// TIA Portal V20 export
// export: Created 2026-10-20T18:54:47.9382926Z, ExportSetting None, DisplayName Totally Integrated Automation Portal, DisplayVersion V20 Update 6, DisplayName TIA Portal Openness, DisplayVersion V20 Update 6, DisplayName TIA Portal Version Control Interface, DisplayVersion V20 Update 6, DisplayName SINAMICS Startdrive Advanced, DisplayVersion V20 SP1, DisplayName SINAMICS Startdrive G130, G150, S120, S150, SINAMICS MV, G220, S200, S210, DisplayVersion V20 SP1, DisplayName SINAMICS Startdrive G110M, G120, G120C, G120D, G120P, G115D, DisplayVersion V20 SP1, DisplayName STEP 7 Professional, DisplayVersion V20 Update 6, DisplayName STEP 7 Safety, DisplayVersion V20 Update 2, DisplayName WinCC Basic/Comfort/Advanced, DisplayVersion V20 Update 6, DisplayName WinCC Unified, DisplayVersion V20 Update 6
VAR_GLOBAL   // PLC tag table "IO_ET200_1"
   "C1102 - SHUTTLE IN POSITION 2" AT %I107.6 : Bool;
   "C1102 - SHUTTLE IN POSITION 1" AT %I107.7 : Bool;
   "C1102 - SENSOR CNV RIGHT (PALLET DETECT 2)" AT %I107.0 : Bool;
   "C1107 - SENSOR CNV LEFT (PALLET DETECT 2)" AT %I127.1 : Bool;
   "C1107 - SHUTTLE IN POSITION 2" AT %I127.6 : Bool;
   "C1107 - SHUTTLE IN POSITION 1" AT %I127.7 : Bool;
   "C1107 - SENSOR CNV RIGHT (PALLET DETECT 2)" AT %I127.0 : Bool;
   "C1107 - SENSOR CNV RIGHT (PALLET DETECT 1)" AT %I127.5 : Bool;
   "C1102 - SENSOR CNV RIGHT (PALLET DETECT 1)" AT %I107.5 : Bool;
   "C1107 - SENSOR CNV LEFT (PALLET DETECT 1)" AT %I126.4 : Bool;
   "C1107 - SENSOR CNV LEFT" AT %I126.5 : Bool;
   "C1106 - SENSOR SAFETY PIN1 DOWN" AT %I115.3 : Bool;
   "C1107 - SENSOR SAFETY PIN1 UP" AT %I127.2 : Bool;
   "C1102 - SENSOR CNV LEFT" AT %I106.5 : Bool;
   "C1102 - SENSOR CNV LEFT (PALLET DETECT 1)" AT %I106.4 : Bool;
   "C1105 - SENSOR SAFETY PIN1 UP" AT %I113.2 : Bool;
   "C1105 - SHUTTLE IN POSITION 2" AT %I113.6 : Bool;
   "C1105 - SHUTTLE IN POSITION 1" AT %I113.7 : Bool;
   "C1105 - SENSOR CNV RIGHT (PALLET DETECT 2)" AT %I113.0 : Bool;
   "C1105 - SENSOR CNV RIGHT (PALLET DETECT 1)" AT %I113.5 : Bool;
   "C1105 - SENSOR CNV LEFT (PALLET DETECT 2)" AT %I113.1 : Bool;
   "C1105 - SENSOR CNV LEFT (PALLET DETECT 1)" AT %I112.4 : Bool;
   "C1105 - SENSOR CNV LEFT" AT %I112.5 : Bool;
   "C1104 - SENSOR SAFETY PIN1 DOWN" AT %I111.3 : Bool;
   "C1104 - SHUTTLE IN POSITION 2" AT %I111.6 : Bool;
   "C1104 - SHUTTLE IN POSITION 1" AT %I111.7 : Bool;
   "C1105 - SENSOR SAFETY PIN1 DOWN" AT %I113.3 : Bool;
   "C1104 - SENSOR CNV RIGHT (PALLET DETECT 2)" AT %I111.0 : Bool;
   "C1104 - SENSOR CNV LEFT (PALLET DETECT 2)" AT %I111.1 : Bool;
   "C1104 - SENSOR CNV LEFT (PALLET DETECT 1)" AT %I110.4 : Bool;
   "C1104 - SENSOR CNV LEFT" AT %I110.5 : Bool;
   "C1104 - SENSOR CNV RIGHT (PALLET DETECT 1)" AT %I111.5 : Bool;
   "C1106 - SENSOR CNV LEFT" AT %I114.5 : Bool;
   "C1106 - SENSOR CNV LEFT (PALLET DETECT 2)" AT %I115.1 : Bool;
   "C1106 - SENSOR CNV LEFT (PALLET DETECT 1)" AT %I114.4 : Bool;
   "C1106 - SENSOR SAFETY PIN1 UP" AT %I115.2 : Bool;
   "C1106 - SHUTTLE IN POSITION 2" AT %I115.6 : Bool;
   "C1106 - SHUTTLE IN POSITION 1" AT %I115.7 : Bool;
   "C1106 - SENSOR CNV RIGHT (PALLET DETECT 2)" AT %I115.0 : Bool;
   "C1106 - SENSOR CNV RIGHT (PALLET DETECT 1)" AT %I115.5 : Bool;
   "C1104 - SENSOR SAFETY PIN1 UP" AT %I111.2 : Bool;
   "C1102 - SENSOR CNV LEFT (PALLET DETECT 2)" AT %I107.1 : Bool;
   "C1107 - SENSOR SAFETY PIN1 DOWN" AT %I127.3 : Bool;
   "C1206 - SENSOR SAFETY PIN1 UP" AT %I345.2 : Bool;
   "C1206 - SHUTTLE IN POSITION 2" AT %I345.6 : Bool;
   "C1206 - SHUTTLE IN POSITION 1" AT %I345.7 : Bool;
   "C1206 - SENSOR CNV RIGHT (PALLET DETECT 2)" AT %I345.1 : Bool;
   "C1206 - SENSOR CNV RIGHT (PALLET DETECT 1)" AT %I344.4 : Bool;
   "C1206 - SENSOR CNV LEFT (PALLET DETECT 2)" AT %I345.0 : Bool;
   "C1206 - SENSOR CNV LEFT (PALLET DETECT 1)" AT %I345.5 : Bool;
   "C1206 - SENSOR CNV LEFT" AT %I345.4 : Bool;
   "C1205 - SENSOR SAFETY PIN1 DOWN" AT %I343.3 : Bool;
   "C1205 - SENSOR SAFETY PIN1 UP" AT %I343.2 : Bool;
   "C1205 - SENSOR CNV RIGHT (PALLET DETECT 2)" AT %I343.1 : Bool;
   "C1205 - SENSOR CNV RIGHT (PALLET DETECT 1)" AT %I342.4 : Bool;
   "C1205 - SENSOR CNV LEFT (PALLET DETECT 2)" AT %I343.0 : Bool;
   "C1205 - SENSOR CNV LEFT (PALLET DETECT 1)" AT %I343.5 : Bool;
   "C1205 - SENSOR CNV LEFT" AT %I343.4 : Bool;
   "C1204 - SENSOR SAFETY PIN1 DOWN" AT %I341.3 : Bool;
   "C1204 - SENSOR SAFETY PIN1 UP" AT %I341.2 : Bool;
   "C1204 - SHUTTLE IN POSITION 1" AT %I341.7 : Bool;
   "C1204 - SENSOR CNV RIGHT (PALLET DETECT 2)" AT %I341.1 : Bool;
   "C1204 - SENSOR CNV RIGHT (PALLET DETECT 1)" AT %I340.6 : Bool;
   "C1206 - SENSOR SAFETY PIN1 DOWN" AT %I345.3 : Bool;
   "C1207 - SENSOR CNV LEFT" AT %I347.4 : Bool;
   "C1207 - SENSOR CNV LEFT (PALLET DETECT 2)" AT %I347.0 : Bool;
   "C1208 - SENSOR CNV RIGHT (PALLET DETECT 1)" AT %I348.4 : Bool;
   "C1207 - SENSOR SAFETY PIN1 DOWN" AT %I347.3 : Bool;
   "C1207 - SENSOR SAFETY PIN1 UP" AT %I347.2 : Bool;
   "C1207 - SHUTTLE IN POSITION 2" AT %I347.6 : Bool;
   "C1207 - SHUTTLE IN POSITION 1" AT %I347.7 : Bool;
   "C1207 - SENSOR CNV RIGHT (PALLET DETECT 2)" AT %I347.1 : Bool;
   "C1207 - SENSOR CNV RIGHT (PALLET DETECT 1)" AT %I346.4 : Bool;
   "C1207 - SENSOR CNV LEFT (PALLET DETECT 1)" AT %I347.5 : Bool;
   "C1204 - SENSOR CNV LEFT (PALLET DETECT 2)" AT %I341.0 : Bool;
   "C1204 - SHUTTLE IN POSITION 2" AT %I341.6 : Bool;
   "C1203 - SENSOR CNV LEFT" AT %I339.4 : Bool;
   "C1203 - SENSOR CNV LEFT (PALLET DETECT 2)" AT %I339.0 : Bool;
   "C1204 - SENSOR CNV LEFT" AT %I341.4 : Bool;
   "C1204 - SENSOR CNV LEFT (PALLET DETECT 1)" AT %I341.5 : Bool;
   "C1203 - SHUTTLE IN POSITION 1" AT %I339.7 : Bool;
   "C1203 - SENSOR CNV RIGHT (PALLET DETECT 2)" AT %I339.1 : Bool;
   "C1203 - SENSOR CNV RIGHT (PALLET DETECT 1)" AT %I338.4 : Bool;
   "C1203 - SHUTTLE IN POSITION 2" AT %I339.6 : Bool;
   "E-STOP L1 - CH1(1)" AT %I528.0 : Bool;
   "E-STOP L1 - CH2(1)" AT %I528.4 : Bool;
   "KEY REMOTE/LOCAL L1 - CH1(1)" AT %I528.1 : Bool;
   "KEY REMOTE/LOCAL L1 - CH2(1)" AT %I528.5 : Bool;
   "C1207 - SENSOR CNV RIGHT" AT %I346.5 : Bool;
   "C1105 - SENSOR CNV RIGHT" AT %I113.4 : Bool;
   "C1106 - SENSOR CNV RIGHT" AT %I115.4 : Bool;
   "C1206 - SENSOR CNV RIGHT" AT %I344.5 : Bool;
   "C1102 - SENSOR CNV RIGHT" AT %I107.4 : Bool;
   "C1104 - SENSOR CNV RIGHT" AT %I111.4 : Bool;
   "C1107 - SENSOR CNV RIGHT" AT %I127.4 : Bool;
   "C1204 - SENSOR CNV RIGHT" AT %I340.7 : Bool;
   "C1205 - SENSOR CNV RIGHT" AT %I342.5 : Bool;
   "C1203 - SENSOR CNV RIGHT" AT %I338.5 : Bool;
   "VTD1 DOCKING PINS RETRACTED 2" AT %I157.3 : Bool;
   "CVTD1 SENSOR CONVEYOR LEFT" AT %I156.1 : Bool;
   "CVTD1 SENSOR CONVEYOR LEFT (PALLET DETECT 1)" AT %I156.2 : Bool;
   "CVTD1 SENSOR CONVEYOR CENTER" AT %I156.0 : Bool;
   "VTD1 DOCKING PINS EXTENDED 1" AT %I157.0 : Bool;
   "C1202 - SHUTTLE IN POSITION 2" AT %I133.6 : Bool;
   "C1202 - SENSOR CNV LEFT (PALLET DETECT 2)" AT %I133.0 : Bool;
   "C1101 - SENSOR CNV LEFT (PALLET DETECT 1)" AT %I104.0 : Bool;   // TESTED
   "C1202 - SENSOR CNV RIGHT" AT %I132.7 : Bool;
   "C1201 - SENSOR CNV LEFT (PALLET DETECT 2)" AT %I131.0 : Bool;   // TESTED
   "C1101 - SHUTTLE IN POSITION 2" AT %I104.2 : Bool;   // TESTED
   "C1101 - SENSOR CNV LEFT (PALLET DETECT 2)" AT %I105.1 : Bool;   // TESTED
   "C1101 - SENSOR CNV RIGHT (PALLET DETECT 2)" AT %I105.0 : Bool;   // TESTED
   "C1201 - SHUTTLE IN POSITION 2" AT %I131.6 : Bool;   // TESTED
   "C1201 - SENSOR CNV RIGHT (PALLET DETECT 1)" AT %I130.4 : Bool;   // TESTED
   "C1201 - SENSOR CNV RIGHT" AT %I130.5 : Bool;   // TESTED
   "C1101 - SENSOR CNV LEFT" AT %I104.1 : Bool;   // TESTED
   "C1101 - SENSOR CNV RIGHT" AT %I104.4 : Bool;   // TESTED
   "C1201 - SENSOR CNV RIGHT (PALLET DETECT 2)" AT %I131.1 : Bool;   // TESTED
   "C1202 - SENSOR CNV LEFT (PALLET DETECT 1)" AT %I133.5 : Bool;
   "C1202 - SENSOR CNV LEFT" AT %I133.4 : Bool;
   "C1202 - SENSOR CNV RIGHT (PALLET DETECT 2)" AT %I133.1 : Bool;
   "C1202 - SENSOR CNV RIGHT (PALLET DETECT 1)" AT %I132.6 : Bool;
   "C1202 - SHUTTLE IN POSITION 1" AT %I133.7 : Bool;
   "C1101 - SHUTTLE IN POSITION 1" AT %I104.3 : Bool;   // TESTED
   "C1201 - SENSOR CNV LEFT" AT %I131.4 : Bool;   // TESTED
   "C1101 - SENSOR CNV RIGHT (PALLET DETECT 1)" AT %I104.5 : Bool;   // TESTED
   "C1201 - SENSOR CNV LEFT (PALLET DETECT 1)" AT %I131.5 : Bool;   // TESTED
   "C1103 - SENSOR CNV LEFT" AT %I108.5 : Bool;
   "C1103 - SENSOR CNV RIGHT (PALLET DETECT 2)" AT %I109.0 : Bool;
   "C1103 - SHUTTLE IN POSITION 2" AT %I109.6 : Bool;
   "C1103 - SENSOR CNV RIGHT" AT %I109.4 : Bool;
   "C1103 - SENSOR CNV LEFT (PALLET DETECT 1)" AT %I108.4 : Bool;
   "C1103 - SENSOR CNV LEFT (PALLET DETECT 2)" AT %I109.1 : Bool;
   "VTD1 DOCKING PINS RETRACTED 1" AT %I157.2 : Bool;
   "VTD1 LEVEL DETECT 1" AT %I157.7 : Bool;
   "VTD1 LEVEL DETECT 2" AT %I157.6 : Bool;
   "VTD1 DOCKING PINS EXTENDED 2" AT %I157.1 : Bool;
   "C1103 - SHUTTLE IN POSITION 1" AT %I109.7 : Bool;
   "C1103 - SENSOR CNV RIGHT (PALLET DETECT 1)" AT %I109.5 : Bool;
   "C1208 - SENSOR SAFETY PIN1 UP" AT %I349.2 : Bool;
   "C1108 - SENSOR SAFETY PIN1 UP" AT %I129.2 : Bool;
   "C1108 - SHUTTLE IN POSITION 2" AT %I129.6 : Bool;
   "C1108 - SHUTTLE IN POSITION 1" AT %I129.7 : Bool;
   "C1208 - SENSOR CNV RIGHT" AT %I348.5 : Bool;
   "C1208 - SENSOR CNV LEFT (PALLET DETECT 2)" AT %I349.0 : Bool;
   "C1201 - SHUTTLE IN POSITION 1" AT %I131.7 : Bool;   // TESTED
   "C1208 - SENSOR CNV RIGHT (PALLET DETECT 2)" AT %I349.1 : Bool;
   "C1208 - SENSOR SAFETY PIN1 DOWN" AT %I349.3 : Bool;
   "C1208 - SHUTTLE IN POSITION 1" AT %I349.7 : Bool;
   "C1108 - SENSOR CNV RIGHT (PALLET DETECT 2)" AT %I129.0 : Bool;
   "C1208 - SHUTTLE IN POSITION 2" AT %I349.6 : Bool;
   "C1208 - SENSOR CNV LEFT" AT %I349.4 : Bool;
   "C1108 - SENSOR CNV LEFT (PALLET DETECT 2)" AT %I129.1 : Bool;
   "C1208 - SENSOR CNV LEFT (PALLET DETECT 1)" AT %I349.5 : Bool;
   "C1108 - SENSOR CNV RIGHT" AT %I129.4 : Bool;
   "C1108 - SENSOR CNV RIGHT (PALLET DETECT 1)" AT %I129.5 : Bool;
   "C1108 - SENSOR CNV LEFT" AT %I128.5 : Bool;
   "C1108 - SENSOR CNV LEFT (PALLET DETECT 1)" AT %I128.4 : Bool;
   "C1108 - SENSOR SAFETY PIN1 DOWN" AT %I129.3 : Bool;
   "VTD1 ULTIMATE SLOWDOWN" AT %I157.4 : Bool;
   "VTD1 ULTIMATE CREEP" AT %I157.5 : Bool;
   "C1102 - SENSOR SAFETY PIN1 UP" AT %I107.2 : Bool;   // TESTED
   "C1102 - SENSOR SAFETY PIN1 DOWN" AT %I107.3 : Bool;   // TESTED
   "C1203 - SENSOR SAFETY PIN1 UP" AT %I339.2 : Bool;   // TESTED
   "C1203 - SENSOR SAFETY PIN1 DOWN" AT %I339.3 : Bool;   // TESTED
   "C1202 - SENSOR SAFETY PIN1 UP" AT %I133.2 : Bool;   // TESTED
   "C1202 - SENSOR SAFETY PIN1 DOWN" AT %I133.3 : Bool;   // 0TESTED
   "E-STOP L7 - CH1(1)" AT %I1179.0 : Bool;
   "KEY REMOTE/LOCAL L6 - CH2(1)" AT %I882.7 : Bool;
   "E-STOP L6 - CH2(1)" AT %I882.6 : Bool;
   "KEY REMOTE/LOCAL L5 - CH2(1)" AT %I882.5 : Bool;
   "E-STOP L5 - CH2(1)" AT %I882.4 : Bool;
   "KEY REMOTE/LOCAL L6 - CH1(1)" AT %I882.3 : Bool;
   "E-STOP L6 - CH1(1)" AT %I882.2 : Bool;
   "KEY REMOTE/LOCAL L5 - CH1(1)" AT %I882.1 : Bool;
   "E-STOP L5 - CH1(1)" AT %I882.0 : Bool;
   "KEY REMOTE/LOCAL L4 - CH2(1)" AT %I636.7 : Bool;
   "KEY REMOTE/LOCAL L7 - CH1(1)" AT %I1179.1 : Bool;
   "E-STOP L4 - CH2(1)" AT %I636.6 : Bool;
   "E-STOP L3 - CH2(1)" AT %I636.4 : Bool;
   "KEY REMOTE/LOCAL L4 - CH1(1)" AT %I636.3 : Bool;
   "E-STOP L4 - CH1(1)" AT %I636.2 : Bool;
   "KEY REMOTE/LOCAL L3 - CH1(1)" AT %I636.1 : Bool;
   "E-STOP L3 - CH1(1)" AT %I636.0 : Bool;
   "KEY REMOTE/LOCAL L2 - CH2(1)" AT %I528.7 : Bool;
   "KEY REMOTE/LOCAL L2 - CH1(1)" AT %I528.3 : Bool;
   "E-STOP L2 - CH2(1)" AT %I528.6 : Bool;
   "E-STOP L2 - CH1(1)" AT %I528.2 : Bool;
   "E-STOP L8 - CH1(1)" AT %I1179.2 : Bool;
   "E-STOP L7 - CH2(1)" AT %I1179.4 : Bool;
   "KEY REMOTE/LOCAL L8 - CH1(1)" AT %I1179.3 : Bool;
   "KEY REMOTE/LOCAL L8 - CH2(1)" AT %I1179.7 : Bool;
   "E-STOP L8 - CH2(1)" AT %I1179.6 : Bool;
   "KEY REMOTE/LOCAL L7 - CH2(1)" AT %I1179.5 : Bool;
   "KEY REMOTE/LOCAL L3 - CH2(1)" AT %I636.5 : Bool;
   "CVTD1 SENSOR CONVEYOR RIGHT (PALLET DETECT 1)" AT %I156.4 : Bool;
   "C1103 - SENSOR SAFETY PIN1 DOWN" AT %I109.3 : Bool;
   "C1103 - SENSOR SAFETY PIN1 UP" AT %I109.2 : Bool;
   "CVTD1 SENSOR CONVEYOR RIGHT" AT %I156.5 : Bool;
   "C1203 - SENSOR CNV LEFT (PALLET DETECT 1)" AT %I339.5 : Bool;
   "C1205 - SHUTTLE IN POSITION 1" AT %I343.7 : Bool;   // DOESN`T HAVE THE MIRROR
   "C1205 - SHUTTLE IN POSITION 2" AT %I343.6 : Bool;   // DOESN`T HAVE THE MIRROR
   "CVTD1 OVERHANG LEFT" AT %I156.7 : Bool;
   "CVTD1 OVERHANG RIGHT" AT %I156.6 : Bool;
END_VAR
